// TIA Portal V20 export
// export: Created 2026-10-12T05:11:21.6829766Z, ExportSetting WithDefaults, DisplayName Totally Integrated Automation Portal, DisplayVersion V20, DisplayName TIA Portal Openness, DisplayVersion V20, DisplayName TIA Portal Teamcenter Gateway, DisplayVersion V20, DisplayName TIA Portal Version Control Interface, DisplayVersion V20, DisplayName SINAMICS Startdrive Advanced, DisplayVersion V20 SP1 Update 2, DisplayName SINAMICS Startdrive G110M, G120, G120C, G120D, G120P, G115D, DisplayVersion V20 SP1 Update 2, DisplayName SINAMICS Startdrive G130, G150, S120, S150, SINAMICS MV, G220, S200, S210, DisplayVersion V20 SP1 Update 2, DisplayName STEP 7 Professional, DisplayVersion V20, DisplayName STEP 7 Safety, DisplayVersion V20, DisplayName WinCC Basic/Comfort/Advanced, DisplayVersion V20, DisplayName WinCC Professional, DisplayVersion V20, DisplayName WinCC Unified, DisplayVersion V20
FUNCTION "FRK_ManualCondition" : Void   // FC82, SCL
{ S7_Optimized_Access := 'TRUE' }
VERSION : 0.1
// stored: AutoNumber true, IsIECCheckEnabled false, SetENOAutomatically false, UDAEnableTagReadback false
   VAR_INPUT
      Slot : Int;
      Value : DInt;
      Ok : Bool;
      Diag : "ST_Diagnostic";
      Bypassable : Bool;
   END_VAR
   VAR_IN_OUT
      Conditions : Array[1..16] of "FRK_ManualConditionRow";
   END_VAR
BEGIN

   IF #Slot < 1 OR #Slot > 16 THEN
       RETURN;
   END_IF;
   #Conditions[#Slot].Used := TRUE;
   #Conditions[#Slot].Value := #Value;
   #Conditions[#Slot].Ok := #Ok;
   #Conditions[#Slot].Diag := #Diag;
   #Conditions[#Slot].Bypassable := #Bypassable;
END_FUNCTION
